(* IEC 61131-3 sources: rungstone/fixtures/plc/iec61499_fill, 2 files *)

(* ---- Fill_61499.st ---- *)
(* GENERATED BY Rungstone - DRAFT FOR ENGINEER REVIEW. Fill_61131.st rewritten for IEC 61499: timers, edges and counters as CYCLE arithmetic. *)
FUNCTION_BLOCK Fill
  VAR_INPUT
    Start_PB : BOOL;
    Level_High : BOOL;
    CYCLE : TIME := T#10ms;
  END_VAR
  VAR_OUTPUT
    Fill_Valve : BOOL;
    Done_Lamp : BOOL;
  END_VAR
  VAR
    Filling : BOOL;
    Fill_Timer_ET : TIME;
    Fill_Timer_Run : BOOL;
    Fill_Timer_Q : BOOL;
    Start_Edge_Mem : BOOL;
    Start_Edge_Q : BOOL;
    Batches_CV : INT;
    Batches_CU_Mem : BOOL;
    Batches_Q : BOOL;
  END_VAR
  (* R_TRIG Start_Edge *)
  Start_Edge_Q := Start_PB AND NOT Start_Edge_Mem;
  Start_Edge_Mem := Start_PB;
  IF Start_Edge_Q THEN Filling := TRUE; END_IF;
  (* TON Fill_Timer: IN = Filling, PT = T#3s *)
  IF Filling THEN
    IF Fill_Timer_Run THEN
      Fill_Timer_ET := Fill_Timer_ET + CYCLE;
      IF Fill_Timer_ET > T#3s THEN Fill_Timer_ET := T#3s; END_IF;
    END_IF;
    Fill_Timer_Run := TRUE;
  ELSE
    Fill_Timer_ET := T#0s;
    Fill_Timer_Run := FALSE;
  END_IF;
  Fill_Timer_Q := Fill_Timer_Run AND Fill_Timer_ET >= T#3s;
  IF Level_High OR Fill_Timer_Q THEN Filling := FALSE; END_IF;
  Fill_Valve := Filling;
  (* CTU Batches: CU = Fill_Timer_Q, PV = 5 *)
  IF Fill_Timer_Q AND NOT Batches_CU_Mem AND Batches_CV < 32767 THEN Batches_CV := Batches_CV + 1; END_IF;
  Batches_CU_Mem := Fill_Timer_Q;
  Batches_Q := Batches_CV >= 5;
  Done_Lamp := Batches_Q;
END_FUNCTION_BLOCK

(* ---- Fill_61131.st ---- *)
(* Scan-style source with TON, R_TRIG and CTU, for the IEC 61499 translation fixture. *)
PROGRAM Fill
  VAR
    Start_PB AT %IX0.0 : BOOL;
    Level_High AT %IX0.1 : BOOL;
    Fill_Valve AT %QX0.0 : BOOL;
    Done_Lamp AT %QX0.1 : BOOL;
  END_VAR
  VAR
    Fill_Timer : TON;
    Start_Edge : R_TRIG;
    Batches : CTU;
    Filling : BOOL;
  END_VAR
  Start_Edge(CLK := Start_PB);
  IF Start_Edge.Q THEN Filling := TRUE; END_IF;
  Fill_Timer(IN := Filling, PT := T#3s);
  IF Level_High OR Fill_Timer.Q THEN Filling := FALSE; END_IF;
  Fill_Valve := Filling;
  Batches(CU := Fill_Timer.Q, RESET := FALSE, PV := 5);
  Done_Lamp := Batches.Q;
END_PROGRAM
